{region 'Documentation'}
(*!
<summary>Captures one snapshot until Reset; Disable/Re-Enable never replaces it.</summary>
<description>

Disabling observation preserves the original snapshot. Re-enabling requires a fresh
preceding observation before comparisons resume; it does not replace that snapshot.

StartIndex is an absolute IN index and Length selects 1..255 elements within IN. Memory
must have at least Length elements from its own lower bound. Invalid references or ranges
report Error.

The caller provides dedicated writable Memory that must not overlap IN; overlap is not
checked. Keep bindings, selected range and snapshot contents stable until Reset. Reset
invalidates the snapshot without clearing Memory bytes.

</description>
*)
{endregion}
FUNCTION_BLOCK AssertArrayNoValueChange_Word EXTENDS AssertionBase
VAR_INPUT
    Mask : WORD := WORD#16#FFFF; //! Bits included in each element comparison.
    StartIndex : DINT; //! First selected index in IN; uses the array's declared index range, not a zero-based offset.
    Length : USINT; //! Number of monitored elements, from 1 through 255.
END_VAR
VAR_IN_OUT CONSTANT
    IN : ARRAY[*] OF WORD; //! Read-only actual data; the selected range must remain stable during the call.
END_VAR
VAR_IN_OUT
    Memory : ARRAY[*] OF WORD; //! Dedicated snapshot storage; only this assertion writes its selected elements.
END_VAR
VAR
    FSnapshotValid : BOOL;
    FObservationPrevious : BOOL;
    FEvaluationActive : BOOL;
END_VAR

SUPER^();

{region 'Documentation'}
(*!
<summary>Capture once or compare against the retained snapshot after range validation.</summary>
*)
{endregion}
METHOD PROTECTED Assert
VAR
    InLowerIndex : DINT;
    InUpperIndex : DINT;
    MemoryLowerIndex : DINT;
    MemoryUpperIndex : DINT;
    MemoryEndIndex : LINT;
    EndIndex : LINT;
    Offset : LINT;
    InIndex : DINT;
    MemoryIndex : DINT;
    Message : STRING(GVL_Constants.MessageLength);
    ReferenceText : STRING(GVL_Constants.AssertionValueLength);
    ActualText : STRING(GVL_Constants.AssertionValueLength);
END_VAR
VAR CONSTANT
    HexDigitCount : USINT := 4;
END_VAR
FEvaluationActive := ObservationActive AND FObservationPrevious AND FSnapshotValid;
FObservationPrevious := ObservationActive;

IF NOT ObservationActive THEN
    RETURN;
END_IF;

IF Result = E_Result.Error THEN
    RETURN;
END_IF;

// C0371: FB inputs are checked here before any reference access.
{warning disable C0371}
IF NOT __ISVALIDREF(IN) THEN
    Error(Message := 'Assertion error: IN reference is invalid.');
    RETURN;
END_IF;

IF NOT __ISVALIDREF(Memory) THEN
    Error(Message := 'Assertion error: Memory reference is invalid.');
    RETURN;
END_IF;

InLowerIndex := LOWER_BOUND(IN, 1);
InUpperIndex := UPPER_BOUND(IN, 1);
MemoryLowerIndex := LOWER_BOUND(Memory, 1);
MemoryUpperIndex := UPPER_BOUND(Memory, 1);
EndIndex := DINT_TO_LINT(StartIndex) + USINT_TO_LINT(Length) - 1;
MemoryEndIndex := DINT_TO_LINT(MemoryLowerIndex) + USINT_TO_LINT(Length) - 1;

IF (Length = 0)
    OR (StartIndex < InLowerIndex) OR (StartIndex > InUpperIndex)
    OR (EndIndex > DINT_TO_LINT(InUpperIndex))
    OR (MemoryEndIndex > DINT_TO_LINT(MemoryUpperIndex)) THEN
    Message := CONCAT('Assertion error: array or memory range is invalid. StartIndex = ',
        DINT_TO_STRING(StartIndex));
    Message := CONCAT(Message, ', EndIndex = ');
    Message := CONCAT(Message, LINT_TO_STRING(EndIndex));
    Message := CONCAT(Message, ', Length = ');
    Message := CONCAT(Message, USINT_TO_STRING(Length));
    Message := CONCAT(Message, '.');
    Error(Message := Message);
    RETURN;
END_IF;

IF NOT FSnapshotValid THEN
    FOR Offset := 0 TO USINT_TO_LINT(Length) - 1 DO
        InIndex := LINT_TO_DINT(DINT_TO_LINT(StartIndex) + Offset);
        MemoryIndex := LINT_TO_DINT(DINT_TO_LINT(MemoryLowerIndex) + Offset);
        Memory[MemoryIndex] := IN[InIndex];
    END_FOR;
    FSnapshotValid := TRUE;
    RETURN;
END_IF;

IF NOT EvaluationActive THEN
    RETURN;
END_IF;

IF Result = E_Result.Failed THEN
    RETURN;
END_IF;

FOR Offset := 0 TO USINT_TO_LINT(Length) - 1 DO
    InIndex := LINT_TO_DINT(DINT_TO_LINT(StartIndex) + Offset);
    MemoryIndex := LINT_TO_DINT(DINT_TO_LINT(MemoryLowerIndex) + Offset);
    IF (IN[InIndex] AND Mask) <> (Memory[MemoryIndex] AND Mask) THEN
        ReferenceText := CreateAssertionTextValue_Hex(Value := WORD_TO_LWORD(Memory[MemoryIndex]),
            DigitCount := HexDigitCount);
        ActualText := CreateAssertionTextValue_Hex(Value := WORD_TO_LWORD(IN[InIndex]),
            DigitCount := HexDigitCount);
        Message := CONCAT('Assertion failed: array value changed. Reference[',
            DINT_TO_STRING(MemoryIndex));
        Message := CONCAT(Message, '] = ');
        Message := CONCAT(Message, ReferenceText);
        Message := CONCAT(Message, ', IN[');
        Message := CONCAT(Message, DINT_TO_STRING(InIndex));
        Message := CONCAT(Message, '] = ');
        Message := CONCAT(Message, ActualText);
        Message := CONCAT(Message, '.');
        Message := CONCAT(Message, ' Mask = ');
        Message := CONCAT(Message, CreateAssertionTextValue_Hex(Value := WORD_TO_LWORD(Mask),
            DigitCount := HexDigitCount));
        Fail(Message := Message);
        RETURN;
    END_IF;
END_FOR;

Pass();
{warning restore C0371}
END_METHOD

{region 'Documentation'}
(*!
<summary>Current/last call has consecutive observation and an existing snapshot.</summary>
*)
{endregion}
{attribute 'monitoring' := 'call'}
PROPERTY PUBLIC EvaluationActive : BOOL //! Current/last call has consecutive observation and an existing snapshot.
GET // PUBLIC
EvaluationActive := FEvaluationActive;
END_GET
END_PROPERTY

{region 'Documentation'}
(*!
<summary>Invalidate the snapshot and observation history.</summary>
<description>

Does not clear external Memory. The next active observation captures a new snapshot
before comparison.

</description>
*)
{endregion}
METHOD PROTECTED ResetAssertion
FSnapshotValid := FALSE;
FObservationPrevious := FALSE;
FEvaluationActive := FALSE;
END_METHOD

END_FUNCTION_BLOCK

(* stored: Version 1.1.0.1
   POU AssertArrayNoValueChange_Word: Id {6f7c23ff-c242-4c01-a4b7-c1d9c135082f}, SpecialFunc None
   Folder Internal: Id {195b962a-29d5-456e-b646-239e90a00621}
   Method Assert: Id {cbf2b9db-e547-4f23-a5e0-8b7662bbf0a9}
   Property EvaluationActive: Id {233520b6-cd95-41b8-ab6c-7d6306046df1}
   Get Get: Id {9468009a-d2df-4e4c-9ce3-f77bbabd00c1}
   Method ResetAssertion: Id {afe7b869-22c1-4d4b-b9fb-199d58aa8854} *)
